SUBAPPLICATION DO_TOGGLE_RPC_QXA_OPC (* Digitaler Freigabe-Ausgang als Klick-Toggle (AX_T_FF_INIT, Default AN): CREATE_METHOD-Server nimmt einen argumentlosen RPC-Trigger von mehreren gleichberechtigten Aufrufern entgegen (z.B. STG1-SoftKey-Relay UND OPC-Dashboard), alle takten denselben CLK - KEIN OR nach dem Flipflop, AX_T_FF_INIT.Q ist alleinige Source of Truth fuer den physischen Ausgang UND den remote publizierten Zustand. Generisch fuer jeden Not-Bedienung-/Strassenmodus-artigen Digital-Toggle-Ausgang mit Mehrfach-Bedienung. *)
  (* Standard: 61499-2 *)
  (* Version 1.4, 2026-11-25, Franz Höpfinger, Meisterschulen am Ostbahnhof, SERVER_0 -> MyLib::net::SERVER_0_QO (IND nur bei QO=TRUE, RSP intern). Ein gescheitertes RSP meldet IND mit QO=FALSE, direkt IND->RSP ergab eine Endlosschleife. *)
  (* Version 1.3, 2026-10-13, Franz Höpfinger, Meisterschulen am Ostbahnhof, Neuer SubAppEventOutput INITO (Type EInit), durchgereicht von DigitalOutput_DO.INITO - analog ILOCK_SWITCH_2_QXA_OPC v1.3, fuer Aufnahme_Option.SUB. *)
  (* Version 1.2, 2026-10-11, Franz Höpfinger, Meisterschulen am Ostbahnhof, Neuer SubAppEventInput INIT (Type EInit), durchgereicht an DigitalOutput_DO.INIT statt Auto-Verteilung - analog ILOCK_SWITCH_2_QXA_OPC v1.2, 'Init wie bei Tecu' (Franz). *)
  (* Version 1.1, 2026-10-11, Franz Höpfinger, Meisterschulen am Ostbahnhof, Neuer QI-InputVar (Default TRUE, rueckwaertskompatibel) durchgereicht an DigitalOutput_DO.QI statt fest verdrahtetem TRUE - analog ILOCK_SWITCH_2_QXA_OPC v1.1. *)
  (* Version 1.0, 2026-09-08, Franz Höpfinger, Meisterschulen am Ostbahnhof, Ausgelagert aus Heben_Senken_TO_QDA_PWM_OPC (Freigabe-DO-Teilnetz) zur Wiederverwendung fuer weitere Digital-Toggle-Ausgaenge. *)
  PACKAGE MyLib::sys;
  IMPORT logiBUS::io::DQ::logiBUS_DO;
  IMPORT logiBUS::io::DQ::logiBUS_DO_S;
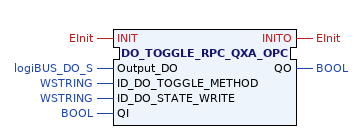
  EVENT_INPUT
    INIT : EInit; (* Initialisierung - vom Aufrufer sequenziert statt per Auto-Verteilung, damit QI vor der physischen Kanalbindung feststeht *)
  END_EVENT
  EVENT_OUTPUT
    INITO : EInit; (* Initialisierung abgeschlossen - echtes Confirm von DigitalOutput_DO.INITO *)
  END_EVENT
  VAR_INPUT
    Output_DO : logiBUS::io::DQ::logiBUS_DO_S := logiBUS_DO::Invalid; (* Physischer Freigabe-Ausgang: Klick-Toggle, Default AN *)
    ID_DO_TOGGLE_METHOD : WSTRING; (* Lokale Methodenadresse (ACTION=CREATE_METHOD) fuer den argumentlosen Freigabe-Toggle-Trigger - wird von mehreren Aufrufern gemeinsam genutzt, alle takten denselben Flipflop *)
    ID_DO_STATE_WRITE : WSTRING; (* Lokale Publish-Adresse (ACTION=WRITE) fuer den tatsaechlichen Freigabe-Zustand (AX_T_FF_INIT.Q) - wird remote abonniert *)
    QI : BOOL := TRUE; (* Qualifier fuer den physischen Ausgang - FALSE haelt diese Instanz komplett inaktiv (keine Hardware-Bindung), fuer den Fall dass derselbe physische Kanal je nach Maschinenvariante anderweitig genutzt wird *)
  END_VAR
  VAR_OUTPUT
    QO : BOOL; (* Quality Output - TRUE if service executed successfully (AND aus DO_TOGGLE_SERVER/AX_T_FF_INIT_DO/PUBLISH_STATE_DO/DigitalOutput_DO) *)
  END_VAR
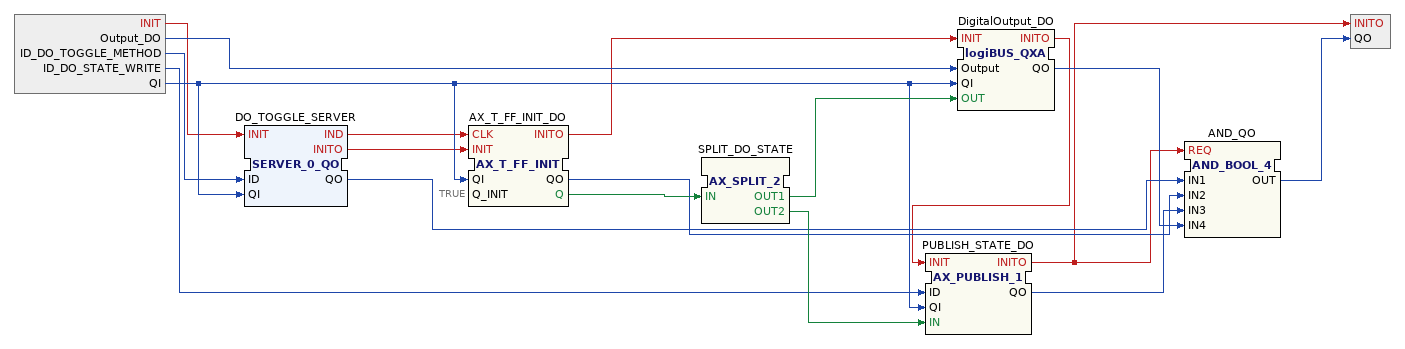
  (* AX_T_FF_INIT.Q ist die EINZIGE Source of Truth fuer DigitalOutput_DO - KEIN AX_OR_2 nach dem Flipflop (anders als TOGGLE_RPC_MERGE_QXA_OPC/Blitzer). Der Methodenaufruf (ID_DO_TOGGLE_METHOD) ist der einzige Eingang und wird von mehreren Aufrufern gemeinsam genutzt - alle takten denselben CLK, kein Merge auf Datenebene noetig. *)
  (* RSP MUSS auf IND zurueckverdrahtet werden (argumentloser Trigger, keine Verarbeitung noetig - wie FORTEs eigener systemtests/clientFailAction.fboot: IND->RSP direkt). Ohne RSP blockiert FORTEs onServerMethodCall den OPC-UA-Server-Thread bis zu 4s (scmMethodCallTimeoutInNanoSeconds) und haelt dabei open62541s globalen serviceMutex - der von JEDEM AX_PUBLISH_1 auf einem anderen FORTE-Thread ebenfalls gebraucht wird. Folge: physischer Ausgang reagiert sofort (kein Lock noetig), aber JEDE OPC-UA-Statusmeldung (nicht nur diese hier) haengt bis zu 4s fest. Siehe Ventilsteuerung/OPC_UA_VERNETZUNG.md Punkt 12. *)
  FBS
    AX_T_FF_INIT_DO : adapter::events::unidirectional::AX_T_FF_INIT(Q_INIT := TRUE);
    SPLIT_DO_STATE : adapter::events::unidirectional::AX_SPLIT_2;
    PUBLISH_STATE_DO : adapter::net::AX_PUBLISH_1;
    DigitalOutput_DO : logiBUS::io::DQ::logiBUS_QXA;
    AND_QO : iec61131::booleanOperators::AND_BOOL_4;
  END_FBS
  SUBAPPS
    DO_TOGGLE_SERVER : MyLib::net::SERVER_0_QO;
  END_SUBAPPS
  EVENT_CONNECTIONS
    DO_TOGGLE_SERVER.IND TO AX_T_FF_INIT_DO.CLK;
    INIT TO DO_TOGGLE_SERVER.INIT;
    DO_TOGGLE_SERVER.INITO TO AX_T_FF_INIT_DO.INIT;
    AX_T_FF_INIT_DO.INITO TO DigitalOutput_DO.INIT;
    PUBLISH_STATE_DO.INITO TO INITO;
    PUBLISH_STATE_DO.INITO TO AND_QO.REQ;
    DigitalOutput_DO.INITO TO PUBLISH_STATE_DO.INIT;
  END_CONNECTIONS
  DATA_CONNECTIONS
    Output_DO TO DigitalOutput_DO.Output;
    QI TO DigitalOutput_DO.QI;
    ID_DO_TOGGLE_METHOD TO DO_TOGGLE_SERVER.ID;
    ID_DO_STATE_WRITE TO PUBLISH_STATE_DO.ID;
    QI TO DO_TOGGLE_SERVER.QI;
    QI TO AX_T_FF_INIT_DO.QI;
    QI TO PUBLISH_STATE_DO.QI;
    DO_TOGGLE_SERVER.QO TO AND_QO.IN1;
    AX_T_FF_INIT_DO.QO TO AND_QO.IN2;
    PUBLISH_STATE_DO.QO TO AND_QO.IN3;
    DigitalOutput_DO.QO TO AND_QO.IN4;
    AND_QO.OUT TO QO;
  END_CONNECTIONS
  ADAPTER_CONNECTIONS
    AX_T_FF_INIT_DO.Q TO SPLIT_DO_STATE.IN;
    SPLIT_DO_STATE.OUT1 TO DigitalOutput_DO.OUT;
    SPLIT_DO_STATE.OUT2 TO PUBLISH_STATE_DO.IN;
  END_CONNECTIONS
END_SUBAPPLICATION
